Universal Robots PolyScope program: JointTargets.urp

Program JointTargets (createdIn=3.0.0 lastSavedIn=3.0.0 directory=/programs installation=default)
Robot Program (runOnlyOnce=true motionType=MoveJ speed=1.047198 acceleration=1.396263 useActiveTCP=false)
  'Program generated by VerticalBot Studio for UR5e on 25/10/2026 12:00:00'
  'Using nominal kinematics.'
  'Using Ref. Frame 2: p[0.100000, -0.050000, 0.020000, 0.000000, 0.000000, 0.523599]'
  'Using TCP Tool 1: p[0.010000, 0.000000, 0.120000, 0.000000, 0.261799, 0.000000]'
  Script: set_tcp(p[0.010000, 0.000000, 0.120000, 0.000000, 0.261799, 0.000000])
  Script: movej([-0.523599, -1.745329, 1.570796, -1.396263, -1.570796, 0.349066],1.20000,0.75000,0,0.0000)
  MoveL speed 250 mm/s, acceleration 1200 mm/s^2 (useActiveTCP=true)
    Waypoint Waypoint_1: position(joints=-0.383972, -1.675516, 1.570796, -1.396263, -1.570796, 0.349066)
  Script: movej([-0.383972, -1.675516, 1.570796, -1.396263, -1.570796, 0.349066],1.20000,0.75000,0,0.0000)
  MoveJ speed 42.97 deg/s, acceleration 68.75 deg/s^2 (useActiveTCP=true)
    Waypoint Waypoint_2: TCP in base x=-441.769 y=44.852 z=400.392 mm, rx=-2.784 ry=-1.254 rz=-0.442 rad; joints [-22, -96, 90, -80, -90, 20] deg; flange x=-456.215 y=40.554 z=519.861 mm, rx=2.8233 ry=1.257 rz=0.075 rad
  MoveL speed 250 mm/s, acceleration 1200 mm/s^2 (useActiveTCP=true)
    Waypoint Waypoint_3: TCP in base x=-415.957 y=97.082 z=429.557 mm, rx=-2.8465 ry=-1.036 rz=-0.3747 rad; joints [-30, -100, 90, -80, -90, 20] deg; flange x=-423.617 y=90.654 z=549.557 mm, rx=2.9521 ry=1.0745 rz=0 rad
    Waypoint Waypoint_4: position(joints=-0.383972, -1.675516, 1.570796, -1.396263, -1.570796, 0.349066)
  Script: movej([-0.523599, -1.745329, 1.570796, -1.396263, -1.570796, 0.349066],1.20000,0.75000,0,0.0000)
  MoveL speed 250 mm/s, acceleration 1200 mm/s^2 (useActiveTCP=true)
    Waypoint Waypoint_5: motionParameters(blendRadius=0.005); position(joints=-0.383972, -1.675516, 1.570796, -1.396263, -1.570796, 0.349066)
  Script: movej([-0.383972, -1.675516, 1.570796, -1.396263, -1.570796, 0.349066],1.20000,0.75000,0,0.0000)
  MoveJ speed 42.97 deg/s, acceleration 68.75 deg/s^2 (useActiveTCP=true)
    Waypoint Waypoint_6: TCP in base x=-441.769 y=44.852 z=400.392 mm, rx=-2.784 ry=-1.254 rz=-0.442 rad; joints [-22, -96, 90, -80, -90, 20] deg; flange x=-456.215 y=40.554 z=519.861 mm, rx=2.8233 ry=1.257 rz=0.075 rad
  MoveL speed 250 mm/s, acceleration 1200 mm/s^2 (useActiveTCP=true)
    Waypoint Waypoint_7: motionParameters(blendRadius=0.005); TCP in base x=-415.957 y=97.082 z=429.557 mm, rx=-2.8465 ry=-1.036 rz=-0.3747 rad; joints [-30, -100, 90, -80, -90, 20] deg; flange x=-423.617 y=90.654 z=549.557 mm, rx=2.9521 ry=1.0745 rz=0 rad
    Waypoint Waypoint_8: motionParameters(blendRadius=0.005); position(joints=-0.383972, -1.675516, 1.570796, -1.396263, -1.570796, 0.349066)
  Script: movej([-0.523599, -1.745329, 1.570796, -1.396263, -1.570796, 0.349066],1.20000,0.75000,0,0.0000)
